(* IEC 61131-3 sources: RAG_PLC/data/result/test/064, 2 files *)

(* ---- wrapped.st ---- *)
(* =========================================================
   Generated by PLC-Eval Benchmark Wrapper
   ========================================================= *)

FUNCTION_BLOCK LLM_Wrapper_FB
VAR_INPUT
    SET : BOOL;
    D0 : BOOL;
    D1 : BOOL;
    D2 : BOOL;
    D3 : BOOL;
    D4 : BOOL;
    D5 : BOOL;
    D6 : BOOL;
    D7 : BOOL;
    CLR : BOOL;
    RST : BOOL;
END_VAR

VAR_OUTPUT
    Q0 : BOOL;
    Q1 : BOOL;
    Q2 : BOOL;
    Q3 : BOOL;
    Q4 : BOOL;
    Q5 : BOOL;
    Q6 : BOOL;
    Q7 : BOOL;
END_VAR

VAR
    edge : BOOL;
END_VAR

IF rst OR set THEN
    Q0 := NOT rst;
    Q1 := Q0;
    Q2 := Q0;
    Q3 := Q0;
    Q4 := Q0;
    Q5 := Q0;
    Q6 := Q0;
    Q7 := Q0;
ELSIF D0 THEN
    Q0 := TRUE;
ELSIF D1 THEN
    Q1 := TRUE;
ELSIF D2 THEN
    Q2 := TRUE;
ELSIF D3 THEN
    Q3 := TRUE;
ELSIF D4 THEN
    Q4 := TRUE;
ELSIF D5 THEN
    Q5 := TRUE;
ELSIF D6 THEN
    Q6 := TRUE;
ELSIF D7 THEN
    Q7 := TRUE;
END_IF;

IF clr AND NOT edge THEN
    IF Q0 THEN
        Q0 := FALSE;
    ELSIF Q1 THEN
        Q1 := FALSE;
    ELSIF Q2 THEN
        Q2 := FALSE;
    ELSIF Q3 THEN
        Q3 := FALSE;
    ELSIF Q4 THEN
        Q4 := FALSE;
    ELSIF Q5 THEN
        Q5 := FALSE;
    ELSIF Q6 THEN
        Q6 := FALSE;
    ELSE
        Q7 := FALSE;
    END_IF;
END_IF;

edge := clr;
END_FUNCTION_BLOCK

PROGRAM Auto_Proxy_Prg
  VAR
    instance : LLM_Wrapper_FB;
  END_VAR

  instance();
END_PROGRAM

CONFIGURATION Config0
  RESOURCE Res0 ON PLC
    TASK TaskMain(INTERVAL := T#20ms, PRIORITY := 0);
    PROGRAM Inst0 WITH TaskMain : Auto_Proxy_Prg;
  END_RESOURCE
END_CONFIGURATION

(* ---- raw_code.st ---- *)
VAR_INPUT
    SET : BOOL;
    D0 : BOOL;
    D1 : BOOL;
    D2 : BOOL;
    D3 : BOOL;
    D4 : BOOL;
    D5 : BOOL;
    D6 : BOOL;
    D7 : BOOL;
    CLR : BOOL;
    RST : BOOL;
END_VAR

VAR_OUTPUT
    Q0 : BOOL;
    Q1 : BOOL;
    Q2 : BOOL;
    Q3 : BOOL;
    Q4 : BOOL;
    Q5 : BOOL;
    Q6 : BOOL;
    Q7 : BOOL;
END_VAR

VAR
    edge : BOOL;
END_VAR

IF rst OR set THEN
    Q0 := NOT rst;
    Q1 := Q0;
    Q2 := Q0;
    Q3 := Q0;
    Q4 := Q0;
    Q5 := Q0;
    Q6 := Q0;
    Q7 := Q0;
ELSIF D0 THEN
    Q0 := TRUE;
ELSIF D1 THEN
    Q1 := TRUE;
ELSIF D2 THEN
    Q2 := TRUE;
ELSIF D3 THEN
    Q3 := TRUE;
ELSIF D4 THEN
    Q4 := TRUE;
ELSIF D5 THEN
    Q5 := TRUE;
ELSIF D6 THEN
    Q6 := TRUE;
ELSIF D7 THEN
    Q7 := TRUE;
END_IF;

IF clr AND NOT edge THEN
    IF Q0 THEN
        Q0 := FALSE;
    ELSIF Q1 THEN
        Q1 := FALSE;
    ELSIF Q2 THEN
        Q2 := FALSE;
    ELSIF Q3 THEN
        Q3 := FALSE;
    ELSIF Q4 THEN
        Q4 := FALSE;
    ELSIF Q5 THEN
        Q5 := FALSE;
    ELSIF Q6 THEN
        Q6 := FALSE;
    ELSE
        Q7 := FALSE;
    END_IF;
END_IF;

edge := clr;
